TYPE ST_EL3351CoeInfo :
STRUCT
	bEnableUserScale: BOOL:= 0;
	diUserScaleOffset: DINT:= 0;
	diUserScaleGain: DINT:= 65536;
	dwFilterSettings: DWORD:= 2;

	bEnableUserScaleIndex8010: BOOL:= 0;
	dnUserScaleOffsetIndex8010: DINT:= 0;
	dnUserScaleGainIndex8010: DINT:= 65536;
END_STRUCT
END_TYPE

(* stored: Version 1.1.0.1, ProductVersion 3.1.4024.15
   DUT ST_EL3351CoeInfo: Id {dcf53909-03c6-4534-b5bd-91672cece6b7} *)
